(* IEC 61131-3 sources: volt/packages/volt-lsp-iec/test-corpus/awa-palletizer/Device/Plc Logic/Application/Library Manager/L_IF1P_FunctionsConnections, 42 files *)

(* ---- L_IF1P_CONNECTDEVICEDATA.dut ---- *)
TYPE L_IF1P_CONNECTDEVICEDATA :
STRUCT
	FUNCTIONMODULEHANDLER : L_IMHP_IModuleHandler;
	DEVICEMODULEHANDLER : L_IMHP_IModuleHandler;
	UISUBDEVICE : UINT := 0;
	EDISCONNECTMODE : L_IF1P_DisconnectMode := L_IF1P_DisconnectMode.Disable;
	SFUNCTIONNAME : STRING;
	SDEVICENAME : STRING;
	ECONNECTIONSTATE : L_IF1P_ConnectionState;
	EERRORID : L_IE1P_Error;
END_STRUCT
END_TYPE

(* ---- L_IF1P_CONNECTEDDEVICEDATA.dut ---- *)
TYPE L_IF1P_CONNECTEDDEVICEDATA :
STRUCT
	FUNCTIONMODULEHANDLER : L_IMHP_IModuleHandler;
	DEVICEMODULEHANDLER : L_IMHP_IModuleHandler;
	SFUNCTIONNAME : STRING;
	UISUBDEVICE : UINT := 0;
	SDEVICENAME : STRING;
	ECONNECTIONSTATE : L_IF1P_ConnectionState;
	EERRORID : L_IE1P_Error;
END_STRUCT
END_TYPE

(* ---- L_IF1P_CONNECTIONINFO.dut ---- *)
TYPE L_IF1P_CONNECTIONINFO :
STRUCT
	PSLAVECONNECTOR : POINTER TO IoConfigConnector;
	UITYPE : UINT;
	UISUBDEVICE : UINT;
	PUTILS : POINTER TO BYTE;
END_STRUCT
END_TYPE

(* ---- L_IF1P_CONNECTIONSTATE.dut ---- *)
TYPE L_IF1P_CONNECTIONSTATE :
(
	UNKNOWN := 0,
	NOTCONNECTED := 1,
	CONNECTING := 2,
	DISCONNECTING := 3,
	CONNECTED := 4,
	ERROR := 10
);
END_TYPE

(* ---- L_IF1P_DISCONNECTDEVICEDATA.dut ---- *)
TYPE L_IF1P_DISCONNECTDEVICEDATA :
STRUCT
	FUNCTIONMODULEHANDLER : L_IMHP_IModuleHandler;
	EMODE : L_IF1P_DisconnectMode := L_IF1P_DisconnectMode.Virtual;
END_STRUCT
END_TYPE

(* ---- L_IF1P_DISCONNECTMODE.dut ---- *)
TYPE L_IF1P_DISCONNECTMODE :
(
	DISABLE := 1,
	VIRTUAL := 2
);
END_TYPE

(* ---- L_IF1P_FUNCITONSINFO.dut ---- *)
TYPE L_IF1P_FUNCITONSINFO :
STRUCT
	PFUNCTIONCONNECTOR : POINTER TO IoConfigConnector;
	UITYPE : UINT;
	ITFFUNCTION : L_IF1P_IFunctionConnection;
END_STRUCT
END_TYPE

(* ---- L_IF1P_INTERNAL.gvl ---- *)
VAR_GLOBAL
	FUNCTIONSTATUSCHANGEDHANDLER : L_IF1P_IConnectionStatusChanged;
	PANYCONNECTOR : POINTER TO IoConfigConnector;
	ITFCONNECTIONHELPER : L_IF1P_IConnectionHelper;
END_VAR

(* ---- L_IF1P_ICONNECTIONHELPER.itf ---- *)
INTERFACE L_IF1P_ICONNECTIONHELPER
END_INTERFACE

METHOD BUILDANDCHECKTABLE
END_METHOD

METHOD FINDCONNECTIONSOURCE : POINTER TO BYTE
VAR_INPUT
	PSLAVECONNECTOR : POINTER TO IoConfigConnector;
	UITYPE : UINT;
	UISUBDEVICE : UINT;
END_VAR
END_METHOD

METHOD FINDFUNCTION : L_IF1P_IFunctionConnection
VAR_INPUT
	PFUNCTIONCONNECTOR : POINTER TO IoConfigConnector;
END_VAR
VAR_OUTPUT
	UITYPE : UINT;
END_VAR
END_METHOD

(* ---- L_IF1P_ICONNECTIONSTATUSCHANGED.itf ---- *)
INTERFACE L_IF1P_ICONNECTIONSTATUSCHANGED
END_INTERFACE

METHOD STATUSCHANGED : BOOL
END_METHOD

(* ---- L_IF1P_IFUNCTIONCONNECTION.itf ---- *)
INTERFACE L_IF1P_IFUNCTIONCONNECTION
END_INTERFACE

METHOD CONNECTDEVICE : UINT
VAR_INPUT
	DEVICEMODULEHANDLER : L_IMHP_IModuleHandler;
	UISUBDEVICE : UINT := 0;
	EDISCONNECTMODE : L_IF1P_DisconnectMode;
	XDISCONNECTEXISTINGCONNECTION : BOOL;
END_VAR
VAR_OUTPUT
	ITFCONNECTIONFBSTATUS : L_IF1P_IStatus;
END_VAR
END_METHOD

METHOD DISCONNECTDEVICE : UINT
VAR_INPUT
	EDISCONNECTMODE : L_IF1P_DisconnectMode;
	XBUSYBEFORE : BOOL;
END_VAR
VAR_OUTPUT
	ITFCONNECTIONFBSTATUS : L_IF1P_IStatus;
END_VAR
END_METHOD

METHOD GEFUNCTIONTINSTANCEPOINTER : POINTER TO BYTE
END_METHOD

METHOD GETCONNECTEDDEVICE : L_IMHP_IModuleHandler
VAR_OUTPUT
	UISUBDEVICE : UINT;
	XVALID : BOOL;
	ITFCONNECTIONFBSTATUS : L_IF1P_IStatus;
END_VAR
END_METHOD

METHOD GETCONNECTIONDIAGNOSTIC
VAR_OUTPUT
	WUSEDBY_COMP : WORD;
	WUSEDBY_SUBCOMP : WORD;
	WACTIVEMODE : WORD;
	WSUBDEVICE : WORD;
	SCONNECTIONSOURE : STRING;
END_VAR
END_METHOD

(* ---- L_IF1P_ISTATUS.itf ---- *)
INTERFACE L_IF1P_ISTATUS
END_INTERFACE

METHOD RESETSTATUS
END_METHOD

(* ---- GETBOOLEANPROPERTY.pou ---- *)
FUNCTION GETBOOLEANPROPERTY : BOOL
VAR_INPUT
	STKEY : WSTRING;
END_VAR
END_FUNCTION

(* ---- GETCOMPANY.pou ---- *)
FUNCTION GETCOMPANY : WSTRING
END_FUNCTION

(* ---- GETNUMBERPROPERTY.pou ---- *)
FUNCTION GETNUMBERPROPERTY : DINT
VAR_INPUT
	STKEY : WSTRING;
END_VAR
END_FUNCTION

(* ---- GETTEXTPROPERTY.pou ---- *)
FUNCTION GETTEXTPROPERTY : WSTRING
VAR_INPUT
	STKEY : WSTRING;
END_VAR
END_FUNCTION

(* ---- GETTEXTPROPERTY2.pou ---- *)
FUNCTION GETTEXTPROPERTY2 : POINTER TO WSTRING
VAR_INPUT
	STKEY : WSTRING;
END_VAR
END_FUNCTION

(* ---- GETTITLE.pou ---- *)
FUNCTION GETTITLE : WSTRING
END_FUNCTION

(* ---- GETVERSION.pou ---- *)
FUNCTION GETVERSION : VERSION
END_FUNCTION

(* ---- GETVERSIONPROPERTY.pou ---- *)
FUNCTION GETVERSIONPROPERTY : VERSION
VAR_INPUT
	STKEY : WSTRING;
END_VAR
END_FUNCTION

(* ---- L_IF1P_CONNECTIONSTATUSCHANGEDEVENT.pou ---- *)
FUNCTION L_IF1P_CONNECTIONSTATUSCHANGEDEVENT : BOOL
END_FUNCTION

(* ---- L_IF1P_FINDCONNECTIONSOURCE.pou ---- *)
FUNCTION L_IF1P_FINDCONNECTIONSOURCE : POINTER TO BYTE
VAR_INPUT
	PSLAVECONNECTOR : POINTER TO IoConfigConnector;
	UITYPE : UINT;
	UISUBDEVICE : UINT;
END_VAR
END_FUNCTION

(* ---- L_IF1P_FINDFUNCTION.pou ---- *)
FUNCTION L_IF1P_FINDFUNCTION : L_IF1P_IFunctionConnection
VAR_INPUT
	PFUNCTIONCONNECTOR : POINTER TO IoConfigConnector;
END_VAR
VAR_OUTPUT
	UITYPE : UINT;
END_VAR
END_FUNCTION

(* ---- L_IF1P_GETIOMGRCONFIGCONNECTORLIST.pou ---- *)
FUNCTION L_IF1P_GETIOMGRCONFIGCONNECTORLIST : RTS_IEC_RESULT
VAR_INPUT
	PPCONNECTORLIST : POINTER TO POINTER TO IoConfigConnector;
	PNCOUNT : POINTER TO DINT;
END_VAR
END_FUNCTION

(* ---- L_IF1P_GETIOMGRCONFIGCOUNTCONNECTOR.pou ---- *)
FUNCTION L_IF1P_GETIOMGRCONFIGCOUNTCONNECTOR : UDINT
VAR_INPUT
	WMODULETYPE : WORD;
END_VAR
END_FUNCTION

(* ---- L_IF1P_GETIOMGRCONFIGFIRSTCHILD.pou ---- *)
FUNCTION L_IF1P_GETIOMGRCONFIGFIRSTCHILD : POINTER TO IoConfigConnector
VAR_INPUT
	PIOCONNECTORLIST : POINTER TO IoConfigConnector;
	PNCOUNT : POINTER TO DINT;
	PFATHER : POINTER TO IoConfigConnector;
END_VAR
END_FUNCTION

(* ---- L_IF1P_GETIOMGRCONFIGGETFIRSTCONNECTOR.pou ---- *)
FUNCTION L_IF1P_GETIOMGRCONFIGGETFIRSTCONNECTOR : POINTER TO IoConfigConnector
VAR_INPUT
	PIOCONNECTORLIST : POINTER TO IoConfigConnector;
	PNCOUNT : POINTER TO DINT;
	WTYPE : WORD;
END_VAR
END_FUNCTION

(* ---- L_IF1P_GETIOMGRCONFIGGETNEXTCONNECTOR.pou ---- *)
FUNCTION L_IF1P_GETIOMGRCONFIGGETNEXTCONNECTOR : POINTER TO IoConfigConnector
VAR_INPUT
	PIOCONNECTORLIST : POINTER TO IoConfigConnector;
	PNCOUNT : POINTER TO DINT;
	WTYPE : WORD;
END_VAR
END_FUNCTION

(* ---- L_IF1P_GETIOMGRCONFIGNEXTCHILD.pou ---- *)
FUNCTION L_IF1P_GETIOMGRCONFIGNEXTCHILD : POINTER TO IoConfigConnector
VAR_INPUT
	PIOCONNECTORLIST : POINTER TO IoConfigConnector;
	PNCOUNT : POINTER TO DINT;
	PFATHER : POINTER TO IoConfigConnector;
END_VAR
END_FUNCTION

(* ---- L_IF1P_GETIOMGRCONFIGPARAMETER.pou ---- *)
FUNCTION L_IF1P_GETIOMGRCONFIGPARAMETER : POINTER TO IoConfigParameter
VAR_INPUT
	PCONNECTOR : POINTER TO IoConfigConnector;
	DWPARAMETERID : DWORD;
END_VAR
END_FUNCTION

(* ---- L_IF1P_GETIOMGRCONFIGPARAMETERVALUEBYTE.pou ---- *)
FUNCTION L_IF1P_GETIOMGRCONFIGPARAMETERVALUEBYTE : BYTE
VAR_INPUT
	PPARAMETER : POINTER TO IoConfigParameter;
	PRESULT : POINTER TO UDINT;
END_VAR
END_FUNCTION

(* ---- L_IF1P_GETIOMGRCONFIGPARAMETERVALUEDWORD.pou ---- *)
FUNCTION L_IF1P_GETIOMGRCONFIGPARAMETERVALUEDWORD : DWORD
VAR_INPUT
	PPARAMETER : POINTER TO IoConfigParameter;
	PRESULT : POINTER TO UDINT;
END_VAR
END_FUNCTION

(* ---- L_IF1P_GETIOMGRCONFIGPARAMETERVALUEWORD.pou ---- *)
FUNCTION L_IF1P_GETIOMGRCONFIGPARAMETERVALUEWORD : WORD
VAR_INPUT
	PPARAMETER : POINTER TO IoConfigParameter;
	PRESULT : POINTER TO UDINT;
END_VAR
END_FUNCTION

(* ---- L_IF1P_INITCONNECTIONTABLEFORSIMULATION.pou ---- *)
FUNCTION L_IF1P_INITCONNECTIONTABLEFORSIMULATION
END_FUNCTION

(* ---- GLOBALTEXTLIST.pou ---- *)
FUNCTION_BLOCK GLOBALTEXTLIST
VAR
	M_TEXTLISTFILE : STRING(255);
	_STNAMESPACE : STRING;
END_VAR
END_FUNCTION_BLOCK

(* ---- L_IF1P_CONNECTDEVICE.pou ---- *)
FUNCTION_BLOCK L_IF1P_CONNECTDEVICE
VAR_INPUT
	XEXECUTE : BOOL;
	FUNCTIONMODULEHANDLER : L_IMHP_IModuleHandler;
	DEVICEMODULEHANDLER : L_IMHP_IModuleHandler;
	UISUBDEVICE : UINT := 0;
	XDISCONNECTEXISTINGCONNECTION : BOOL := TRUE;
	EDISCONNECTMODE : L_IF1P_DisconnectMode := L_IF1P_DisconnectMode.Disable;
END_VAR
VAR_OUTPUT
	XBUSY : BOOL;
	XDONE : BOOL;
	XERROR : BOOL;
	EERRORID : L_IE1P_Error;
END_VAR
VAR
	PDEVICECONNECTOR : POINTER TO IOconfigConnector;
	PFUNCTIONCONNECTOR : POINTER TO IOconfigConnector;
	ITFFUNCTION : L_IF1P_IFunctionConnection;
	UITYPE : UINT;
	XEXECUTEOLD : BOOL;
	FUNCTIONMODULEHANDLEROLD : L_IMHP_IModuleHandler;
	DEVICEMODULEHANDLEROLD : L_IMHP_IModuleHandler;
	SFUNCTIONNAME : STRING;
	SDEVICENAME : STRING;
	ITFCONNECTSTATUS : L_IF1P_IStatus;
	XACTIVE : BOOL;
	ERROR_FUNCTIONMODULEINVALID : WORD := 26001;
	ERROR_DEVICEMODULEINVALID : WORD := 26002;
	ERROR_FUNCTIONMODULENOTSUPPORTED : WORD := 26003;
	ERROR_DEVICEMODULENOTSUPPORTED : WORD := 26004;
	ERROR_NOTSUPPORTEDBYMODULEHANDLERVERSION : WORD := 26005;
	ERROR_INVALIDDISCONNECTMODE : WORD := 26006;
END_VAR
END_FUNCTION_BLOCK

(* ---- L_IF1P_DEVICECONNECTIONHANDLER.pou ---- *)
FUNCTION_BLOCK L_IF1P_DEVICECONNECTIONHANDLER
VAR_INPUT
	XEXECUTE : BOOL;
	ASCCONNECTIONDATA : POINTER TO L_IF1P_ConnectDeviceData;
	XDISCONNECTEXISTINGCONNECTION : BOOL := TRUE;
END_VAR
VAR_OUTPUT
	XBUSY : BOOL;
	XDONE : BOOL;
	XERROR : BOOL;
	EERRORID : L_IE1P_Error;
END_VAR
VAR
	UITYPE : UINT;
	XEXECUTEOLD : BOOL;
	UIIDX : DINT;
	FB_CONNECTDEVICE : L_IF1P_ConnectDevice;
	FB_DISCONNECTDEVICE : L_IF1P_DisconnectDevice;
	XBUSYINTERNAL : BOOL;
	XERRORINTERNAL : BOOL;
	XDONEINTERNAL : BOOL;
	EERRORIDINTERNAL : L_IE1P_Error;
	XCOLLECTINGERROR : BOOL;
	EERRORIDTMP : L_IE1P_Error;
END_VAR
END_FUNCTION_BLOCK

METHOD GETCONNECTIONSTATE : L_IF1P_ConnectionState
VAR_OUTPUT
	EERRORID : L_IE1P_Error;
END_VAR
END_METHOD

METHOD RESET
END_METHOD

(* ---- L_IF1P_DISCONNECTDEVICE.pou ---- *)
FUNCTION_BLOCK L_IF1P_DISCONNECTDEVICE
VAR_INPUT
	XEXECUTE : BOOL;
	FUNCTIONMODULEHANDLER : L_IMHP_IModuleHandler;
	EDISCONNECTMODE : L_IF1P_DisconnectMode := L_IF1P_DisconnectMode.Disable;
END_VAR
VAR_OUTPUT
	XBUSY : BOOL;
	XDONE : BOOL;
	XERROR : BOOL;
	EERRORID : L_IE1P_Error;
END_VAR
VAR
	PDEVICECONNECTOR : POINTER TO IOconfigConnector;
	PFUNCTIONCONNECTOR : POINTER TO IOconfigConnector;
	ITFFUNCTION : L_IF1P_IFunctionConnection;
	UITYPE : UINT;
	XEXECUTEOLD : BOOL;
	FUNCTIONMODULEHANDLEROLD : L_IMHP_IModuleHandler;
	SFUNCTIONNAME : STRING;
	ITFCONNECTIONSTATUS : L_IF1P_IStatus;
	XACTIVE : BOOL;
	ERROR_FUNCTIONMODULEINVALID : WORD := 26001;
	ERROR_DEVICEMODULEINVALID : WORD := 26002;
	ERROR_FUNCTIONMODULENOTSUPPORTED : WORD := 26003;
	ERROR_DEVICEMODULENOTSUPPORTED : WORD := 26004;
	ERROR_NOTSUPPORTEDBYMODULEHANDLERVERSION : WORD := 26005;
	ERROR_INVALIDDISCONNECTMODE : WORD := 26006;
END_VAR
END_FUNCTION_BLOCK

(* ---- L_IF1P_FUNCTIONCONNECTIONVIEWER.pou ---- *)
FUNCTION_BLOCK L_IF1P_FUNCTIONCONNECTIONVIEWER EXTENDS IoDrvBase
VAR
	M_IIODRV : ICmpIoDrv;
	M_IIODRVPARAMETER : ICmpIoDrvParameter;
	DWDISPLAYSELCMD : DWORD;
	BYREQUESTID : BYTE;
	WPAROFFSET : WORD;
	XVALIDAXISSTRING : BOOL;
	SCONNECTEDAXIS1 : STRING;
	SCONNECTEDAXIS2 : STRING;
	DWSTATUSCHANGED : DWORD;
	WRITEPARACOUNT : DWORD;
	CONNECTCOUNT : DWORD;
	READPARACOUNT1 : DWORD;
	READPARACOUNT2 : DWORD;
	READPARACOUNT3 : DWORD;
	WVERSIONMODE : WORD := 0;
	UDICOUNTDEV : UDINT;
	UDICOUNTFUN : UDINT;
	PDATADEVICES : POINTER TO ARRAY [0..255] OF L_IF1P_ConnectionInfo;
	PDATAFUNCTIONS : POINTER TO ARRAY [0..255] OF L_IF1P_FuncitonsInfo;
	HEVENTDOWNLOADDONE : RTS_IEC_HANDLE;
	HINTERFACEDOWNLOADDONE : RTS_IEC_HANDLE;
	HEVENTRESETDONE : RTS_IEC_HANDLE;
	HINTERFACERESETDONE : RTS_IEC_HANDLE;
	ITFCALLBACK : CmpEventMgr.ICmpEventCallback;
	XCONFIGDONE : BOOL;
	XCONFIGBUSY : BOOL;
	WCONFIGCALL : WORD;
	SCOMNAME_DEVICES : STRING := 'Connection_Devices';
	SCOMNAME_FUNCTIONS : STRING := 'Connection_Funcitons';
END_VAR
END_FUNCTION_BLOCK

METHOD BUILDANDCHECKTABLE
END_METHOD

METHOD BUILDUPCONNECTIONTABLE : BOOL
END_METHOD

METHOD FINDCONNECTIONSOURCE : POINTER TO BYTE
VAR_INPUT
	PSLAVECONNECTOR : POINTER TO IoConfigConnector;
	UITYPE : UINT;
	UISUBDEVICE : UINT;
END_VAR
END_METHOD

METHOD FINDFUNCTION : L_IF1P_IFunctionConnection
VAR_INPUT
	PFUNCTIONCONNECTOR : POINTER TO IoConfigConnector;
END_VAR
VAR_OUTPUT
	UITYPE : UINT;
END_VAR
END_METHOD

METHOD GETCONNECTEDSLAVE : BOOL
END_METHOD

METHOD INITIALIZE : UDINT
VAR_INPUT
	WMODULETYPE : UINT;
	DWINSTANCE : UDINT;
	PCONNECTOR : POINTER TO IoConfigConnector;
END_VAR
END_METHOD

METHOD IODRVREADPARAMETER : UDINT
VAR_INPUT
	PCONNECTOR : POINTER TO IoConfigConnector;
	PPARAMETER : POINTER TO IoConfigParameter;
	PDATA : POINTER TO BYTE;
	DWBITSIZE : DWORD;
	DWBITOFFSET : DWORD;
END_VAR
END_METHOD

METHOD IODRVUPDATECONFIGURATION : UDINT
VAR_INPUT
	PCONNECTORLIST : POINTER TO IoConfigConnector;
	NCOUNT : DINT;
END_VAR
END_METHOD

METHOD IODRVUPDATEMAPPING : UDINT
VAR_INPUT
	PTASKMAPLIST : POINTER TO IoConfigTaskMap;
	NCOUNT : DINT;
END_VAR
END_METHOD

METHOD IODRVWRITEPARAMETER : UDINT
VAR_INPUT
	PCONNECTOR : POINTER TO IoConfigConnector;
	PPARAMETER : POINTER TO IoConfigParameter;
	PDATA : POINTER TO BYTE;
	DWBITSIZE : DWORD;
	DWBITOFFSET : DWORD;
END_VAR
END_METHOD

METHOD QUERYINTERFACE : POINTER TO POINTER TO BYTE
VAR_INPUT
	IID : DWORD;
	PRESULT : POINTER TO UDINT;
END_VAR
END_METHOD

METHOD STATUSCHANGED : BOOL
END_METHOD

METHOD FB_EXIT : BOOL
VAR_INPUT
	BINCOPYCODE : BOOL;
END_VAR
END_METHOD

METHOD FB_INIT : BOOL
VAR_INPUT
	BINITRETAINS : BOOL;
	BINCOPYCODE : BOOL;
END_VAR
END_METHOD

METHOD EVENTCALLBACK : UDINT
VAR_INPUT
	PEVENTPARAM : POINTER TO EventParam;
END_VAR
END_METHOD

METHOD REGISTEREVENT
END_METHOD

METHOD UNREGISTEREVENT
END_METHOD

(* ---- L_IF1P_GETCONNECTEDDEVICE.pou ---- *)
FUNCTION_BLOCK L_IF1P_GETCONNECTEDDEVICE
VAR_INPUT
	XEXECUTE : BOOL;
	FUNCTIONMODULEHANDLER : L_IMHP_IModuleHandler;
END_VAR
VAR_OUTPUT
	XBUSY : BOOL;
	XDONE : BOOL;
	XERROR : BOOL;
	EERRORID : L_IE1P_Error;
	ECONNECTIONSTATE : L_IF1P_ConnectionState;
	DEVICEMODULEHANDLER : L_IMHP_IModuleHandler;
	UISUBDEVICE : UINT := 0;
	SDEVICENAME : STRING;
END_VAR
VAR
	PDEVICECONNECTOR : POINTER TO IOconfigConnector;
	PFUNCTIONCONNECTOR : POINTER TO IOconfigConnector;
	ITFFUNCTION : L_IF1P_IFunctionConnection;
	UITYPE : UINT;
	XEXECUTEOLD : BOOL;
	FUNCTIONMODULEHANDLEROLD : L_IMHP_IModuleHandler;
	SFUNCTIONNAME : STRING;
	XVALID : BOOL;
	ITFCONNECTIONSTATUS : L_IF1P_IStatus;
	XACTIVE : BOOL;
	ERROR_FUNCTIONMODULEINVALID : WORD := 26001;
	ERROR_DEVICEMODULEINVALID : WORD := 26002;
	ERROR_FUNCTIONMODULENOTSUPPORTED : WORD := 26003;
	ERROR_DEVICEMODULENOTSUPPORTED : WORD := 26004;
	ERROR_NOTSUPPORTEDBYMODULEHANDLERVERSION : WORD := 26005;
	ERROR_INVALIDDISCONNECTMODE : WORD := 26006;
END_VAR
END_FUNCTION_BLOCK

(* ---- L_IF1P_GETCONNECTEDDEVICES.pou ---- *)
FUNCTION_BLOCK L_IF1P_GETCONNECTEDDEVICES
VAR_INPUT
	XEXECUTE : BOOL;
	ASCCONNECTEDDEVICEDATA : POINTER TO L_IF1P_ConnectedDeviceData;
END_VAR
VAR_OUTPUT
	XBUSY : BOOL;
	XDONE : BOOL;
	XERROR : BOOL;
	EERRORID : L_IE1P_Error;
END_VAR
VAR
	ITFFUNCTION : L_IF1P_IFunctionConnection;
	UITYPE : UINT;
	XEXECUTEOLD : BOOL;
	DIIDX : DINT;
	FB_GETCONNECTEDDEVICE : L_IF1P_GetConnectedDevice;
	SIZE : DINT;
	AVISUDATAARRAY : ARRAY [0..4] OF L_IF1P_ConnectedDeviceData;
	DIACTVALUE : DINT;
	DIMAXVALUE : DINT := 0;
	CDIMINVALUE : DINT := 0;
END_VAR
END_FUNCTION_BLOCK

METHOD UPDATEVISU
END_METHOD

(* ---- L_IF1P_STATUS.pou ---- *)
FUNCTION_BLOCK L_IF1P_STATUS
VAR
	XBUSY : BOOL;
	XDONE : BOOL;
	XERROR : BOOL;
	EERRORID : L_IE1P_Error;
	BUSY : BOOL;
	DONE : BOOL;
	ERROR : BOOL;
	ERRORID : L_IE1P_Error;
END_VAR
END_FUNCTION_BLOCK

METHOD RESETSTATUS
END_METHOD

METHOD SETBUSYSTATE
END_METHOD

METHOD SETDONESTATE : BOOL
END_METHOD

METHOD SETERRORSTATE : BOOL
VAR_INPUT
	ERRORID : L_IE1P_Error;
END_VAR
END_METHOD
